Universal Robots PolyScope program: SetProg.urp

Program SetProg (createdIn=3.0.0 lastSavedIn=3.0.0 directory=/programs installation=default)
Robot Program (runOnlyOnce=true motionType=MoveJ speed=1.047198 acceleration=1.396263 useActiveTCP=false)
  'Program generated by RoboDK v6.0.7 for ABB IRB 120-3/0.6 on XX/XX/XXXX 18:00:00'
  'Using nominal kinematics.'
  'Using Ref. Frame S: p[1.234570, -0.098765, 0.050500, 0.000000, 0.000000, 0.523599]'
  'Using TCP Tool S: p[0.010000, 0.020000, 0.150000, 0.000000, 0.000000, 0.000000]'
  Script: set_tcp(p[0.010000, 0.020000, 0.150000, 0.000000, 0.000000, 0.000000])
  Script: movej([0.000000, -0.174533, 0.349066, 0.000000, 0.523599, 0.000000],1.20000,0.75000,0,0.0000)
  MoveJ speed 42.97 deg/s, acceleration 68.75 deg/s^2 (useActiveTCP=true)
    Waypoint Waypoint_1: TCP in base x=426.318 y=20 z=422.034 mm, rx=0 ry=2.2689 rz=0 rad; joints [0, -10, 20, 0, 30, 0] deg; flange x=317.839 y=0 z=526.113 mm, rx=0 ry=2.2689 rz=0 rad
  MoveL speed 250 mm/s, acceleration 1200 mm/s^2 (useActiveTCP=true)
    Waypoint Waypoint_2: position(joints=0.000000, -0.174533, 0.349066, 0.000000, 0.523599, 0.000000)
  'Circular movement using joint targets is not supported. Change the target type to cartesian or use a joint movement.'
  Script: movej([0.349066, -0.174533, 0.349066, 0.000000, 0.523599, 0.000000],1.20000,0.75000,0,0.0000)
  Wait Sleep waitTime=0.25
  Script: movej([0.523599, -0.349066, 0.698132, 1.047198, -0.785398, -1.745329],1.20000,0.75000,0,0.0000)
  MoveJ speed 42.97 deg/s, acceleration 68.75 deg/s^2 (useActiveTCP=true)
    Waypoint Waypoint_3: TCP in base x=408.367 y=83.8 z=505.12 mm, rx=-0.4874 ry=1.4458 rz=-0.7473 rad; joints [30, -20, 40, 60, -45, -100] deg; flange x=257.546 y=97.782 z=512.713 mm, rx=-0.4874 ry=1.4458 rz=-0.7473 rad
